{attribute 'Tc2GvlVarNames'}
VAR_CONFIG
END_VAR
VAR_CONFIG
	MAIN.Axis.PlcToNc AT %QB0: PLCTONC_AXIS_REF;
	MAIN.Axis.NcToPlc AT %IB0 : NCTOPLC_AXIS_REF;
END_VAR

(* stored: Version 1.1.0.1, ProductVersion 3.1.4024.16
   GVL Variable_Configuration: Id {4da002c0-56e5-454c-b388-02436cb26103} *)
